RESOURCE RES0 : EMB_RES_ECO
  FBS
    DPAC_FULLINIT1 : DPAC_FULLINIT;
    AGUA_REUSO : Agua_Reuso(cfgTempoBoia := 10, cfgBoiaInvertida := FALSE, cfgTempoCom := 5);
    SUB_R1_A6_DI32K0 : IO_DI32(WORD0 := '$${PATH}SUB_R1_A6_DI32K_WORD0', WORD1 := '$${PATH}SUB_R1_A6_DI32K_WORD1', CONN := '$${PATH}SUB_R1_CONN', FALHA_COM := 'RES0.AGUA_REUSO.stsFalhaRemota1', DI_9 := 'RES0.AGUA_REUSO.stsBoiaLSL', DI_0 := 'RES0.DosagemAlcalinizante.BO_800_02.stsSemFalha', DI_1 := 'RES0.DosagemAlcalinizante.DO_800_04.stsLocal', DI_2 := 'RES0.DosagemAlcalinizante.DO_800_04.stsRemoto', DI_3 := 'RES0.DosagemAlcalinizante.DO_800_04.stsLigado', DI_4 := 'RES0.DosagemAlcalinizante.DO_800_04.stsSemFalha', DI_5 := 'RES0.DosagemAlcalinizante.DO_800_05.stsLocal', DI_6 := 'RES0.DosagemAlcalinizante.DO_800_05.stsRemoto', DI_7 := 'RES0.DosagemAlcalinizante.DO_800_05.stsLigado', DI_8 := 'RES0.DosagemAlcalinizante.DO_800_05.stsSemFalha');
    SUBESTACAO : Subestacao(cfgTempoDiscordancia := 5, cfgTempoComGerador := 10, cfgTempoPulsoDisjuntor := 1, cfgTempoRespostaDisjuntor := 5);
    SUB_R1_A3_DI32K0 : IO_DI32(WORD0 := '$${PATH}SUB_R1_A3_DI32K_WORD0', WORD1 := '$${PATH}SUB_R1_A3_DI32K_WORD1', CONN := 'RES0.SUB_R1_A6_DI32K0.SUB_R1_CONN', FALHA_COM := 'RES0.SUBESTACAO.stsFalhaRemota1', DI_0 := 'RES0.SUBESTACAO.djPCE_SUBESTACAO', DI_1 := 'RES0.Pre_Tratamento1.BombaGordura.stsLocal', DI_2 := 'RES0.Pre_Tratamento1.BombaGordura.stsRemoto', DI_3 := 'RES0.Pre_Tratamento1.BombaGordura.stsLigado', DI_4 := 'RES0.Pre_Tratamento1.BombaGordura.stsSemFalha', DI_5 := 'RES0.Pre_Tratamento1.BombaGordura.stsProtecaoTermica', DI_18 := 'RES0.SUBESTACAO.djV4603', DI_19 := 'RES0.SUBESTACAO.djV4604', DI_20 := 'RES0.SUBESTACAO.djCOMP_500_02', DI_21 := 'RES0.SUBESTACAO.djUCT_200_01', DI_22 := 'RES0.SUBESTACAO.djPCM_EEE_BRUTO', DI_23 := 'RES0.SUBESTACAO.djQGBT_220V', DI_24 := 'RES0.SUBESTACAO.djPCM_DESINFECCAO', DI_25 := 'RES0.SUBESTACAO.djBANCO_CAPACITORES', DI_26 := 'RES0.SUBESTACAO.djRES_A1', DI_27 := 'RES0.SUBESTACAO.djRES_A2', DI_28 := 'RES0.SUBESTACAO.mpL_1q1', DI_29 := 'RES0.SUBESTACAO.mpR_1q1', DI_30 := 'RES0.SUBESTACAO.mpP_1q1', DI_31 := 'RES0.SUBESTACAO.mpC_1q1');
    SUB_R1_A4_DI32K0 : IO_DI32(WORD0 := '$${PATH}SUB_R1_A4_DI32K_WORD0', WORD1 := '$${PATH}SUB_R1_A4_DI32K_WORD1', CONN := 'RES0.SUB_R1_A6_DI32K0.SUB_R1_CONN', DI_0 := 'RES0.SUBESTACAO.mpSF_1q1', DI_1 := 'RES0.SUBESTACAO.mpAB_1q1', DI_2 := 'RES0.SUBESTACAO.mpFE_1q1', DI_3 := 'RES0.SUBESTACAO.mpL_1q0', DI_4 := 'RES0.SUBESTACAO.mpR_1q0', DI_5 := 'RES0.SUBESTACAO.mpP_1q0', DI_6 := 'RES0.SUBESTACAO.mpC_1q0', DI_7 := 'RES0.SUBESTACAO.mpSF_1q0', DI_8 := 'RES0.SUBESTACAO.mpAB_1q0', DI_9 := 'RES0.SUBESTACAO.mpFE_1q0', DI_10 := 'RES0.SUBESTACAO.mpL_1q2', DI_11 := 'RES0.SUBESTACAO.mpR_1q2', DI_12 := 'RES0.SUBESTACAO.mpP_1q2', DI_13 := 'RES0.SUBESTACAO.mpC_1q2', DI_14 := 'RES0.SUBESTACAO.mpSF_1q2', DI_15 := 'RES0.SUBESTACAO.mpAB_1q2', DI_16 := 'RES0.SUBESTACAO.mpFE_1q2', DI_17 := 'RES0.Pre_Tratamento2.BombaGordura.stsLocal', DI_18 := 'RES0.Pre_Tratamento2.BombaGordura.stsRemoto', DI_19 := 'RES0.Pre_Tratamento2.BombaGordura.stsLigado', DI_20 := 'RES0.Pre_Tratamento2.BombaGordura.stsSemFalha', DI_21 := 'RES0.Pre_Tratamento2.BombaGordura.stsProtecaoTermica', DI_30 := 'RES0.SUBESTACAO.djV4601', DI_31 := 'RES0.SUBESTACAO.djV4602');
    SUB_R1_A5_DI32K0 : IO_DI32(WORD0 := '$${PATH}SUB_R1_A5_DI32K_WORD0', WORD1 := '$${PATH}SUB_R1_A5_DI32K_WORD1', CONN := 'RES0.SUB_R1_A6_DI32K0.SUB_R1_CONN', DI_0 := 'RES0.SUBESTACAO.djCOMP_500_01', DI_1 := 'RES0.SUBESTACAO.djUCT_200_02', DI_2 := 'RES0.SUBESTACAO.djUCT_200_03', DI_3 := 'RES0.SUBESTACAO.djPCM_NEREDA', DI_4 := 'RES0.SUBESTACAO.djPCM_LODO', DI_5 := 'RES0.SUBESTACAO.djCAP2', DI_6 := 'RES0.SUBESTACAO.djPCM_AGUA_REUSO', DI_7 := 'RES0.SUBESTACAO.djMO_500_01', DI_8 := 'RES0.SUBESTACAO.djRES_B1', DI_9 := 'RES0.SUBESTACAO.djRES_B2', DI_10 := 'RES0.SUBESTACAO.djRES_B3', DI_11 := 'RES0.SUBESTACAO.djQGBT_220V_ENTRADA', DI_12 := 'RES0.SUBESTACAO.djQL_ADM', DI_13 := 'RES0.SUBESTACAO.djQL_PORTARIA', DI_14 := 'RES0.SUBESTACAO.djQLSL', DI_15 := 'RES0.SUBESTACAO.djQL_ILUMINACAO', DI_16 := 'RES0.SUBESTACAO.djPCE_SOPRADORES', DI_17 := 'RES0.SUBESTACAO.djQL_LODO', DI_18 := 'RES0.SUBESTACAO.djRES_C1', DI_19 := 'RES0.SUBESTACAO.djRES_C2', DI_20 := 'RES0.SUBESTACAO.djRES_C3', DI_21 := 'RES0.SUBESTACAO.djRES_C4', DI_22 := 'RES0.SUBESTACAO.djRES_C5', DI_23 := 'RES0.SUBESTACAO.djRES_C6');
    SUB_R1_A8_DQ32K0 : IO_DQ32(WORD0 := '$${PATH}SUB_R1_A8_DQ32K_WORD0', WORD1 := '$${PATH}SUB_R1_A8_DQ32K_WORD1_NAO_USADA', CONN := 'RES0.SUB_R1_A6_DI32K0.SUB_R1_CONN', DO_0 := 'RES0.Pre_Tratamento1.BombaGordura.cmdAcionamento', DO_1 := 'RES0.Pre_Tratamento1.BombaGordura.cmdReset', DO_5 := 'RES0.SUBESTACAO.cmdAbrir1q1', DO_6 := 'RES0.SUBESTACAO.cmdFechar1q1', DO_7 := 'RES0.SUBESTACAO.cmdAbrir1q0', DO_8 := 'RES0.SUBESTACAO.cmdFechar1q0', DO_9 := 'RES0.SUBESTACAO.cmdAbrir1q2', DO_10 := 'RES0.SUBESTACAO.cmdFechar1q2', DO_11 := 'RES0.Pre_Tratamento2.BombaGordura.cmdAcionamento', DO_12 := 'RES0.Pre_Tratamento2.BombaGordura.cmdReset', DO_15 := 'RES0.DosagemAlcalinizante.BO_800_02.cmdAcionamento');
    MGE_AGUA_REUSO : MGE_Generico(cfgTempoCom := 5);
    MGE_QGBT_220V : MGE_Generico(cfgTempoCom := 5);
    Pre_Tratamento1 : UCT_PreTratamento(cfgInstalada := TRUE, cfgTempoCom := 10, cfgTempoReset := 2);
    Pre_Tratamento2 : UCT_PreTratamento(cfgInstalada := TRUE, cfgTempoCom := 10, cfgTempoReset := 2);
    Pre_Tratamento3 : UCT_PreTratamento(cfgInstalada := FALSE, cfgTempoCom := 10, cfgTempoReset := 2);
    FT_40_02 : Sensor_Generico(cfgComunicacao := FALSE, cfgNivel := FALSE, cfgBrutoMin := 4000.0, cfgBrutoMax := 20000.0, cfgFalhaMin := 3800.0, cfgFalhaMax := 22000.0, cfgTempoFalha := 5, cfgUsaConexao := TRUE, cfgUnidade := 'm3/h', cfgCasasDecimais := 1);
    EEEB_A2_DI32K0 : IO_DI32(WORD0 := '$${PATH}EEEB_A2_DI32K_WORD0', WORD1 := '$${PATH}EEEB_A2_DI32K_WORD1', CONN := '$${PATH}EEEB_A2_DI32K0_CONN', DI_1 := 'RES0.EEEB.stsEmergenciaPainel', DI_12 := 'RES0.EEEB.BS_100_01.stsLocal', DI_13 := 'RES0.EEEB.BS_100_01.stsRemoto', DI_14 := 'RES0.EEEB.BS_100_01.stsLigado', DI_15 := 'RES0.EEEB.BS_100_01.stsSemFalha', DI_16 := 'RES0.EEEB.BS_100_01.stsProtecaoTermica', DI_17 := 'RES0.EEEB.BS_100_02.stsLocal', DI_18 := 'RES0.EEEB.BS_100_02.stsRemoto', DI_19 := 'RES0.EEEB.BS_100_02.stsLigado', DI_20 := 'RES0.EEEB.BS_100_02.stsSemFalha', DI_21 := 'RES0.EEEB.BS_100_02.stsProtecaoTermica', DI_22 := 'RES0.EEEB.BS_100_03.stsLocal', DI_23 := 'RES0.EEEB.BS_100_03.stsRemoto', DI_24 := 'RES0.EEEB.BS_100_03.stsLigado', DI_25 := 'RES0.EEEB.BS_100_03.stsSemFalha', DI_26 := 'RES0.EEEB.BS_100_03.stsProtecaoTermica', DI_27 := 'RES0.EEEB.stsBoiaNivelBaixo', DI_28 := 'RES0.EEEB.stsBoiaNivelAlto');
    EEEB_A3_DQ32TK0 : IO_DQ32(WORD0 := '$${PATH}EEEB_A3_DQ32TK_WORD0', WORD1 := '$${PATH}EEEB_A3_DQ32TK_WORD1', CONN := 'RES0.EEEB_A2_DI32K0.EEEB_A2_DI32K0_CONN', DO_0 := 'RES0.EEEB.BS_100_01.cmdAcionamento', DO_1 := 'RES0.EEEB.BS_100_01.cmdReset', DO_2 := 'RES0.EEEB.BS_100_02.cmdAcionamento', DO_3 := 'RES0.EEEB.BS_100_02.cmdReset', DO_4 := 'RES0.EEEB.BS_100_03.cmdAcionamento', DO_5 := 'RES0.EEEB.BS_100_03.cmdReset');
    EEEB : EEE_Bruto(geradorConectado := TRUE, cfgTempoFalhaBoiaL := 10, cfgTempoPartidaPressao := 30, cfgUsaFalhaComunicacao := TRUE);
    MGE_EEE_BRUTO : MGE_Generico(cfgTempoCom := 5);
    SUBNER_A3_DI32K0 : IO_DI32(WORD0 := '$${PATH}SUBNER_A3_DI32K_WORD0', WORD1 := '$${PATH}SUBNER_A3_DI32K_WORD1', CONN := '$${PATH}SUBNER_CONN', FALHA_COM := 'RES0.SUBESTACAO.stsFalhaRemotaNER', DI_0 := 'RES0.SUBESTACAO.djNER_PCE', DI_2 := 'RES0.SUBESTACAO.djNER_PCM', DI_6 := 'RES0.SUBESTACAO.djMO_300_01', DI_22 := 'RES0.SUBESTACAO.djR4005A', DI_23 := 'RES0.SUBESTACAO.djR4005B');
    SUBNER_A4_DI32K0 : IO_DI32(WORD0 := '$${PATH}SUBNER_A4_DI32K_WORD0', WORD1 := '$${PATH}SUBNER_A4_DI32K_WORD1', CONN := 'RES0.SUBNER_A3_DI32K0.SUBNER_CONN', DI_2 := 'RES0.SUBESTACAO.djP4901', DI_3 := 'RES0.SUBESTACAO.djP4902', DI_4 := 'RES0.SUBESTACAO.djP4903');
    SUBEEEB_A2_DI32K0 : IO_DI32(WORD0 := '$${PATH}SUBEEEB_A2_DI32K_WORD0', WORD1 := '$${PATH}SUBEEEB_A2_DI32K_WORD1', CONN := '$${PATH}SUBEEEB_CONN', FALHA_COM := 'RES0.SUBESTACAO.stsFalhaRemotaEEEB', DI_0 := 'RES0.SUBESTACAO.djEEEB_PCE', DI_2 := 'RES0.SUBESTACAO.djEEEB_PCM', DI_6 := 'RES0.SUBESTACAO.djCO_100_01', DI_7 := 'RES0.SUBESTACAO.djCO_100_02', DI_8 := 'RES0.SUBESTACAO.djCO_100_03', DI_9 := 'RES0.SUBESTACAO.djCO_100_04', DI_10 := 'RES0.SUBESTACAO.djGM_100_01_02', DI_11 := 'RES0.SUBESTACAO.djMO_100_01');
    SUBDES_A2_DI32K0 : IO_DI32(WORD0 := '$${PATH}SUBDES_A2_DI32K_WORD0', WORD1 := '$${PATH}SUBDES_A2_DI32K_WORD1', CONN := '$${PATH}SUBDES_CONN', FALHA_COM := 'RES0.SUBESTACAO.stsFalhaRemotaDES', DI_0 := 'RES0.SUBESTACAO.djDES_PCE_DESLIGADO', DI_1 := 'RES0.SUBESTACAO.djDES_PCM_DESLIGADO', DI_2 := 'RES0.SUBESTACAO.djUV_700_01', DI_3 := 'RES0.SUBESTACAO.djUV_700_02', DI_4 := 'RES0.SUBESTACAO.djVC_700_01', DI_5 := 'RES0.SUBESTACAO.djMO_700_01');
    SUBLODO_A3_DI32K0 : IO_DI32(WORD0 := '$${PATH}SUBLODO_A3_DI32K_WORD0', WORD1 := '$${PATH}SUBLODO_A3_DI32K_WORD1', CONN := '$${PATH}SUBLODO_CONN', FALHA_COM := 'RES0.SUBESTACAO.stsFalhaRemotaLODO', DI_0 := 'RES0.SUBESTACAO.dj900_PCE_DESL', DI_2 := 'RES0.SUBESTACAO.dj900_PCM', DI_3 := 'RES0.SUBESTACAO.dj900_SO_01', DI_8 := 'RES0.SUBESTACAO.dj900_SO_02', DI_13 := 'RES0.SUBESTACAO.dj900_AD_01', DI_14 := 'RES0.SUBESTACAO.dj900_AD_02', DI_15 := 'RES0.SUBESTACAO.dj900_AD_03', DI_16 := 'RES0.SUBESTACAO.dj900_PP_01', DI_17 := 'RES0.SUBESTACAO.dj900_MN_01', DI_18 := 'RES0.SUBESTACAO.dj900_MN_02', DI_19 := 'RES0.SUBESTACAO.dj900_MN_03', DI_20 := 'RES0.SUBESTACAO.dj900_MN_04', DI_21 := 'RES0.SUBESTACAO.dj900_MN_05', DI_22 := 'RES0.SUBESTACAO.dj900_BO_01', DI_28 := 'RES0.SUBESTACAO.dj900_BO_02');
    SUBLODO_A4_DI32K0 : IO_DI32(WORD0 := '$${PATH}SUBLODO_A4_DI32K_WORD0', WORD1 := '$${PATH}SUBLODO_A4_DI32K_WORD1', CONN := 'RES0.SUBLODO_A3_DI32K0.SUBLODO_CONN', DI_2 := 'RES0.SUBESTACAO.dj900_BO_03', DI_8 := 'RES0.SUBESTACAO.dj900_BR_01', DI_14 := 'RES0.SUBESTACAO.dj900_BR_02', DI_20 := 'RES0.SUBESTACAO.dj900_VA_01', DI_21 := 'RES0.SUBESTACAO.dj900_VA_02', DI_22 := 'RES0.SUBESTACAO.dj900_VE_01', DI_23 := 'RES0.SUBESTACAO.dj900_VE_02', DI_25 := 'RES0.SUBESTACAO.dj900_VA_06', DI_26 := 'RES0.SUBESTACAO.dj900_VA_07', DI_27 := 'RES0.SUBESTACAO.dj900_VA_08', DI_28 := 'RES0.SUBESTACAO.dj900_VA_09', DI_29 := 'RES0.SUBESTACAO.dj900_VA_10', DI_30 := 'RES0.SUBESTACAO.dj900_VA_11', DI_31 := 'RES0.SUBESTACAO.dj900_VA_12');
    SUBLODO_A5_DI32K0 : IO_DI32(WORD0 := '$${PATH}SUBLODO_A5_DI32K_WORD0', WORD1 := '$${PATH}SUBLODO_A5_DI32K_WORD1', CONN := 'RES0.SUBLODO_A3_DI32K0.SUBLODO_CONN', DI_0 := 'RES0.SUBESTACAO.dj900_VA_13', DI_1 := 'RES0.SUBESTACAO.dj900_VB_03', DI_2 := 'RES0.SUBESTACAO.dj900_VB_04');
    Gradeamento : Gradeamento_Inovaisa;
    DosagemAlcalinizante : Dosagem_Alcalinizante;
    SR_SUB_R1_REMOTA1 : Status_Remota;
    SR_SUB_R2_REMOTA2 : Status_Remota;
    SR_SUB_NER_REMOTA1 : Status_Remota;
    SR_NER_R2_FT02 : Status_Remota;
    SR_EEEB_A1_REMOTA : Status_Remota;
    SR_SUB_EEEB_REMOTA : Status_Remota;
    SR_SUB_DESINF_REMOTA : Status_Remota;
  END_FBS
  EVENT_CONNECTIONS
    SUBESTACAO.921BB7D26016F39E TO Pre_Tratamento1.0B595E2D755381E4;
    SUBESTACAO.921BB7D26016F39E TO Pre_Tratamento2.0B595E2D755381E4;
    SUBESTACAO.921BB7D26016F39E TO Pre_Tratamento3.0B595E2D755381E4;
    Pre_Tratamento1.5A6CC858EDC95420 TO Pre_Tratamento2.0B595E2D755381E4;
    Pre_Tratamento2.5A6CC858EDC95420 TO Pre_Tratamento3.0B595E2D755381E4;
    SUBESTACAO.921BB7D26016F39E TO DosagemAlcalinizante.3550FA6DB34A3727;
    SUBESTACAO.921BB7D26016F39E TO Gradeamento.D1B66AFAEC6D2FF0;
    START.COLD TO DPAC_FULLINIT1.INIT;
    START.WARM TO DPAC_FULLINIT1.INIT;
    START.ONLINECHANGE TO DPAC_FULLINIT1.OC_RETRIGGER;
  END_CONNECTIONS
  DATA_CONNECTIONS
    SUBESTACAO.FEF1963C61B73419 TO Pre_Tratamento1.2C19134423AEFFAA;
    SUBESTACAO.FEF1963C61B73419 TO Pre_Tratamento2.2C19134423AEFFAA;
    SUBESTACAO.FEF1963C61B73419 TO Pre_Tratamento3.2C19134423AEFFAA;
    SUBESTACAO.5DB035BC4F7321F6 TO Pre_Tratamento1.D205F407BC981FB4;
    SUBESTACAO.E3892FBEADB0545B TO Pre_Tratamento2.D205F407BC981FB4;
    SUBESTACAO.85B535DFB1FB677D TO Pre_Tratamento3.D205F407BC981FB4;
    Pre_Tratamento1.1F8CA54F12D8796B TO Pre_Tratamento2.3F3598C544A33E47;
    Pre_Tratamento1.A737D1113B918FC6 TO Pre_Tratamento2.BFB78C58CA08F906;
    Pre_Tratamento2.1F8CA54F12D8796B TO Pre_Tratamento3.3F3598C544A33E47;
    Pre_Tratamento2.A737D1113B918FC6 TO Pre_Tratamento3.BFB78C58CA08F906;
    SUBESTACAO.B9F74BEEB26000F4 TO DosagemAlcalinizante.A0398C4E77A10EEE;
    SUBESTACAO.499BDAC4EA9F62DF TO DosagemAlcalinizante.7CA01E1D24150792;
    SUBESTACAO.FEF1963C61B73419 TO DosagemAlcalinizante.7838A99D6B60D295;
    SUBESTACAO.2BBFC35BA4EC9BC5 TO Gradeamento.358F3774D14189DB;
    SUBESTACAO.FEF1963C61B73419 TO Gradeamento.98A20843E1C25CF2;
  END_CONNECTIONS
END_RESOURCE
